Fanuc KAREL source: KT00529.KL

PROGRAM KT00529
%NOLOCKGROUP
VAR
  P1: XYZWPREXT
  P2: JOINTPOS
  OUT: POSITION
BEGIN
  P1.X = 1.0
  OUT = P1 : P2
END KT00529
